// TIA Portal V20 export
// export: Created 2026-10-12T15:46:51.766989Z, ExportSetting WithDefaults, DisplayName Totally Integrated Automation Portal, DisplayVersion V20, DisplayName TIA Portal Openness, DisplayVersion V20, DisplayName TIA Portal Teamcenter Gateway, DisplayVersion V20, DisplayName TIA Portal Version Control Interface, DisplayVersion V20, DisplayName SINAMICS Startdrive Advanced, DisplayVersion V20 SP1 Update 2, DisplayName SINAMICS Startdrive G110M, G120, G120C, G120D, G120P, G115D, DisplayVersion V20 SP1 Update 2, DisplayName SINAMICS Startdrive G130, G150, S120, S150, SINAMICS MV, G220, S200, S210, DisplayVersion V20 SP1 Update 2, DisplayName STEP 7 Professional, DisplayVersion V20, DisplayName STEP 7 Safety, DisplayVersion V20, DisplayName WinCC Basic/Comfort/Advanced, DisplayVersion V20, DisplayName WinCC Professional, DisplayVersion V20, DisplayName WinCC Unified, DisplayVersion V20
FUNCTION "FRK_JsonRecord" : Bool   // FC128, SCL
{ S7_Optimized_Access := 'TRUE' }
VERSION : 0.1
// stored: AutoNumber true, IsIECCheckEnabled false, SetENOAutomatically false, UDAEnableTagReadback false
   VAR_INPUT
      Data : "ST_ConfigRecord";
   END_VAR
   VAR_IN_OUT
      Line : WString;
   END_VAR
   VAR_TEMP
      Ok : Bool;
      Flag : WString[1];
   END_VAR
BEGIN

   #FRK_JsonRecord := FALSE;
   #Line := WSTRING#'{';
   #Ok := "FRK_JsonAdd"(Key := 'scope', Value := STRING_TO_WSTRING(#Data.Scope), Quoted := TRUE, LastField := FALSE, Line := #Line);
   IF NOT #Ok THEN
       #Line := WSTRING#'';
       RETURN;
   END_IF;
   #Ok := "FRK_JsonAdd"(Key := 'key', Value := STRING_TO_WSTRING(#Data.WriteKey), Quoted := TRUE, LastField := FALSE, Line := #Line);
   IF NOT #Ok THEN
       #Line := WSTRING#'';
       RETURN;
   END_IF;
   #Ok := "FRK_JsonAdd"(Key := 'rev', Value := UDINT_TO_WSTRING(#Data.Revision), Quoted := FALSE, LastField := FALSE, Line := #Line);
   IF NOT #Ok THEN
       #Line := WSTRING#'';
       RETURN;
   END_IF;
   #Ok := "FRK_JsonAdd"(Key := 'kind', Value := DINT_TO_WSTRING(#Data.Kind), Quoted := FALSE, LastField := FALSE, Line := #Line);
   IF NOT #Ok THEN
       #Line := WSTRING#'';
       RETURN;
   END_IF;
   #Ok := "FRK_JsonAdd"(Key := 'type', Value := DINT_TO_WSTRING(#Data.ValueType), Quoted := FALSE, LastField := FALSE, Line := #Line);
   IF NOT #Ok THEN
       #Line := WSTRING#'';
       RETURN;
   END_IF;
   #Ok := "FRK_JsonAdd"(Key := 'value', Value := STRING_TO_WSTRING(#Data.ValueText), Quoted := TRUE, LastField := TRUE, Line := #Line);
   IF NOT #Ok THEN
       #Line := WSTRING#'';
       RETURN;
   END_IF;
   #FRK_JsonRecord := TRUE;
END_FUNCTION
